FUNCTION_BLOCK EPUCK_INIT (* E-puck initialization *)
  (* Standard: 61499-2; Classification: SIFB; ApplicationDomain: Robotics; Function: Robot initialization; Type: SIFB; Description: Initialize e-puck1 motors and sensors *)
  (* Version 1.0, 2026-10-22, Mauricio Martins Taques Filho, GASR/UDESC, Initial version *)
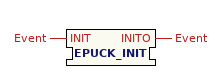
  EVENT_INPUT
    INIT; (* Robot initialization *)
  END_EVENT
  EVENT_OUTPUT
    INITO; (* Robot ready *)
  END_EVENT
  SERVICE APPLICATION/RESOURCE
    SEQUENCE Initialization
      APPLICATION.INIT() -> APPLICATION.INITO();
    END_SEQUENCE
  END_SERVICE
END_FUNCTION_BLOCK
